// TEST DI F_TimeToSeconds E F_SecondsToTime
FUNCTION_BLOCK FB_Conversion_Test EXTENDS TcUnit.FB_TestSuite
VAR
END_VAR

TimeToSeconds();
SecondsToTime();

METHOD PRIVATE SecondsToTime
TEST('SecondsToTime');

AssertEquals_TIME(
	Expected	:=	T#2S250MS,
	Actual		:=	ML.F_SecondsToTime(2.25),
	Message		:=	'2,25 s');

TEST_FINISHED();
END_METHOD

METHOD PRIVATE TimeToSeconds
TEST('TimeToSeconds');

AssertEquals_REAL(
	Expected	:=	1.5,
	Actual		:=	ML.F_TimeToSeconds(T#1S500MS),
	Delta		:=	0.0001,
	Message		:=	'1,5 s');

TEST_FINISHED();
END_METHOD

END_FUNCTION_BLOCK

(* stored: Version 1.1.0.1, ProductVersion 3.1.4024.9
   POU FB_Conversion_Test: Id {9598820b-4ec5-4366-bc8e-dcb57e3e867a}, SpecialFunc None
   Folder METHODs: Id {781ef806-dbbf-4156-973a-77174c7fb02d}
   Method SecondsToTime: Id {1a5bf50d-42af-455b-82fe-89ee347ff27b}
   Method TimeToSeconds: Id {141153eb-4b2f-4d65-88ac-1ba507bc60f2} *)
